Staubli VAL3: CalToolPos4.pgx

public program CalToolPos4(tool& x_tTool)
  local bool l_bStatus
  local pointRx l_p1
  local pointRx l_p2
  local pointRx l_p3
  local pointRx l_p4
  local point l_pCenter
  local tool l_t1
  local tool l_t2
  local tool l_t3
  local tool l_t4
  local num x1
  local num x2
  local num x3
  local num x4
  local num y1
  local num y2
  local num y3
  local num y4
  local num z1
  local num z2
  local num z3
  local num z4
begin
  //取中心点xyz
  l_p1=db:pTeach1
  l_p2=db:pTeach2
  l_p3=db:pTeach3
  l_p4=db:pTeach4
  l_pCenter=here(flange,world)
  call _CalpSphere(l_p1,l_p2,l_p3,l_p4,l_pCenter,l_bStatus)

  if l_bStatus==false
    call db:hmiAlert("DeviationIsTooLarge","warning")
  else
    if db:sMounting=="Floor"
      l_pCenter.trsf.rx=0
      l_pCenter.trsf.ry=180
      l_pCenter.trsf.rz=0
    elseIf db:sMounting=="Ceiling"
      l_pCenter.trsf.rx=0
      l_pCenter.trsf.ry=0
      l_pCenter.trsf.rz=0
    endIf
    l_t1.trsf=!l_p1.trsf*l_pCenter.trsf
    l_t2.trsf=!l_p2.trsf*l_pCenter.trsf
    l_t3.trsf=!l_p3.trsf*l_pCenter.trsf
    l_t4.trsf=!l_p4.trsf*l_pCenter.trsf
    x_tTool.trsf.x=(l_t1.trsf.x+l_t2.trsf.x+l_t3.trsf.x+l_t4.trsf.x)/4
    x_tTool.trsf.y=(l_t1.trsf.y+l_t2.trsf.y+l_t3.trsf.y+l_t4.trsf.y)/4
    x_tTool.trsf.z=(l_t1.trsf.z+l_t2.trsf.z+l_t3.trsf.z+l_t4.trsf.z)/4
    x_tTool.trsf.rx=l_t1.trsf.rx
    x_tTool.trsf.ry=l_t1.trsf.ry
    x_tTool.trsf.rz=l_t1.trsf.rz
    call db:hmiAlert("SaveInTool1","info")
  endIf
end
